(* IEC 61131-3 sources: daoli-st-library/DL_Motion (part 25) *)

(* ---- FB_DL_ToolChangerSeq.st ---- *)
(*
    FB_DL_ToolChangerSeq —— 换刀机构顺控（刀位校验 → 取刀 → 换刀 → 旧刀回库 → 到位确认）
    ------------------------------------------------------------------
    组件名称  : FB_DL_ToolChangerSeq
    分类      : DL_Motion / ToolChange
    前缀      : FB_DL_
    版本      : 1.0.0
    溯源      : 借鉴组织 —— T2-6 Rockwell AOI（矩阵行 166，伺服外围件方向）
                + 次源 t1-9 国产机床 FB 手册公开功能清单（换刀必有反馈对与
                互锁为公开工程惯例）；clean-room 声明 —— 状态机 / 码位 /
                时序 100% 自有，零代码行复制，无闭源参考。
    平台      : 纯 IEC 61131-3（ENUM + CASE + TON / R_TRIG），CODESYS 3.5 /
                TwinCAT 3 / InoProShop / Machine Expert 通用
    作者      : 道莅代码库 · PLC编程专家（R72 构建轮 · 批 4 · 序号 10）
    ------------------------------------------------------------------
    功能说明  : 换刀机构「命令 - 反馈 - 确认」编排：eIdle → eSelect（刀位
                校验 / 映射，发刀位指令，等刀库对位与机械手原位）→ ePick
                （机械手取刀，正向反馈对）→ eSwap（主轴换刀，bSpindleFree
                互锁迁入，反向反馈对）→ eReturn（旧刀回库，回原位反馈）→
                eDone（bToolDone 单拍脉冲）→ eIdle。每执行相带独立超时
                （单 TON 实例，PT = tActTimeout，相驻留即 IN，R145 相级
                看门狗口径），超时 → eFault + 锁存码。
                受理语义（同拍竞态闸，R279）：换刀受理只看 uToolReq **值
                变更沿**的迁入沿锁存副本 _uReqLatch，运行中禁跨拍双判——
                运行中刀位号变更被忽略（沿已被消费），须再次变更刀位号
                （或先归 0）才重新受理；同值重发须先归 0 或变更刀位号
                （接口契约声明，无执行沿引脚的替代口径）。
                安全语义：
                ① eSwap 为安全相，迁入必带全量闸位复检（bSpindleFree +
                   NOT _bFault，R274）；
                ② 换刀中途 bSpindleFree 撤销 → **保持相 + 信息提示，不中断
                   不回退**（防半程掉刀，安全侧声明；继续完成换刀比半程
                   悬臂更安全）；
                ③ 失能 / 故障 → 全输出清零 + 状态回 eIdle（停机相输出清零，
                   R57）；失能不清故障锁存（操作态非复位），复位沿才解除；
                ④ uToolReq = 0 或 > nToolCount → 拒收 + 信息码，不发任何
                   指令；nToolCount = 1（单刀库退化）→ 信息级直接
                   eSelect→ePick（跳过刀库对位等待）。
    错误码    : 16#0004_08B0 刀位请求越域（0 或 > nToolCount），已拒收不发
                            指令 —— 信息级，不置 bError（R45）
                16#0004_08B1 单刀库退化（nToolCount = 1），eSelect 直接转
                            ePick —— 信息级，不置 bError
                16#0004_08B2 执行相超时（任一执行相驻留超 tActTimeout），
                            锁存至复位沿 —— 故障级
                16#0004_08B3 换刀相主轴互锁撤销（bSpindleFree 于 eSwap 内
                            为 FALSE），保持相照走 —— 信息级，不置 bError
                16#0004_08B4 组态非法（nToolCount = 0 / tActTimeout 非正），
                            锁存至复位沿 —— 故障级
                加码反证句（R90）：08B2 / 08B4 输出同为 eFault + bError，
                但 08B4 在 eIdle 即锁存（无执行史）、08B2 必有执行相驻留史
                （eState 轨迹可证），成因互斥不可互换观测；08B0 / 08B1 /
                08B3 各有独立触发事件（拒收沿 / 组态相 / 互锁撤销拍），
                不由现有输出组合还原，故各立一码。
    码位总账  : 16#0004_08B0 用 ｜ 16#0004_08B1 用 ｜ 16#0004_08B2 用 ｜
                16#0004_08B3 用 ｜ 16#0004_08B4 用
                （08A6 / 08A7 已由 FB_DL_TurretToolSelect 占用，本件不占）
    边界与披露: 一 R_TRIG（rtReq / rtReset）与 TON（tonAct）每拍**无条件
                   调用**（规则 ⑦）；tonAct IN = 执行相驻留判据显式变量
                   （R145 看门狗使能只用相驻留，不叠业务条件补集）；超时
                   判定在 CASE 之后（本拍完成事件优先，R275 同拍竞态口径），
                   超时有一拍检测延迟（声明口径）；
                二 零全局变量、零 VAR_EXTERNAL、零物理地址；
                三 归属 Ownership：E_DL_ToolChangePhase 属主为本文件（全库
                   唯一定义，R264），引用件只引用不重声明；
                四 状态机 ENUM + CASE 必带 ELSE 兜底（非法枚举值 → eFault
                   锁存）；段 5b 统一故障迁入闸（R274 迁入完备性）；
                五 反馈引脚语义声明：bToolHome = 所选刀位对位取刀口、
                   bArmHome = 机械手原位、bArmFwd = 机械臂正向到位、
                   bArmBack = 机械臂反向到位，均引脚注入，本件不发轴指令；
                六 分工声明：FB_DL_TurretToolSelect（刀塔分度就近选刀解算，
                   无机械手取放编排）、FB_DL_ToolLifeBudget（寿命记账）——
                   本件只管换刀机构「命令 - 反馈 - 确认」时序编排，刀位
                   就近解算归刀塔件、寿命记账归记账件，互引不互代；
                七 依赖声明：仅 Standard.library（TON / R_TRIG），零厂商
                   方言；
                八 复位沿作用域（R311 逐项声明）：清故障锁存 + 清锁存码 +
                   迁 eIdle + 清 _uReqPrev（强制下次刀位值变更沿可受理），
                   **不清**周期计数类（本件无）与 _uReqLatch（回 Idle 后由
                   下次受理沿重写）。
    验收向量  : V1 正常换刀（uToolReq = 3，nToolCount = 8，反馈按时序到）
                → eState 轨迹 eIdle→eSelect→ePick→eSwap→eReturn→eDone→
                eIdle，bToolDone 单拍，eFault 不出现；
                V2 uToolReq = 0 → 08B0 拒收不发指令；V3 nToolCount = 1 →
                08B1 + eSelect 直转 ePick；V4 eSwap 中 bSpindleFree 撤销
                → 保持相照走 + 08B3；V5 任一执行相超时 → 08B2 锁存 +
                eFault + 输出清零；V6 复位沿 → 解锁回 eIdle；
                V7 nToolCount = 0 → 08B4 锁存；V8 失能 → 输出清零 +
                eIdle，锁存保留。
                算法已证（脚本）：未跑 ｜ 编译器已证（三平台）：未跑
    修订记录  : 2026-11-23 v1.0.0 首次入库（R72 构建轮 · 批 4 · 序号 10）
*)
TYPE E_DL_ToolChangePhase :
(
    eIdle   := 0,                          // 空闲：等刀位请求值变更沿 / idle, waiting for a tool request change edge
    eSelect := 10,                         // 刀位校验：发刀位指令，等刀库对位与机械手原位 / select, issue the tool command
    ePick   := 20,                         // 取刀：机械臂正向，等正向到位 / pick, the arm forward to the magazine
    eSwap   := 30,                         // 换刀：主轴互锁迁入，机械臂反向 / swap, gated by the spindle free interlock
    eReturn := 40,                         // 旧刀回库：机械臂正向回原位 / return, the old tool back to the magazine
    eDone   := 50,                         // 完成：bToolDone 单拍脉冲相 / done, the one shot pulse phase
    eFault  := 60                          // 故障：锁存待复位 / fault, latched until the reset
);
END_TYPE

FUNCTION_BLOCK FB_DL_ToolChangerSeq
VAR_INPUT
    uToolReq     : UINT := 0;              (* 目标刀位请求，[刀位]，1 起计，0 或越容量拒收 / the requested tool number, refused when zero or over capacity *)
    nToolCount   : UINT := 8;              (* 刀库容量组态，[刀位]，禁 0 / the magazine tool count, must not be zero *)
    bToolHome    : BOOL := FALSE;          (* 所选刀位对位反馈，[标志]，引脚注入 / the tool position aligned feedback *)
    bArmHome     : BOOL := FALSE;          (* 机械手原位反馈，[标志]，引脚注入 / the arm home feedback *)
    bArmFwd      : BOOL := FALSE;          (* 机械臂正向到位反馈，[标志]，引脚注入 / the arm forward in position feedback *)
    bArmBack     : BOOL := FALSE;          (* 机械臂反向到位反馈，[标志]，引脚注入 / the arm backward in position feedback *)
    bSpindleFree : BOOL := FALSE;          (* 主轴可换刀互锁，[标志]，eSwap 迁入与驻留判据 / the spindle free interlock *)
    tActTimeout  : TIME := T#10S;          (* 执行相超时，[ms]，禁非正 / the action phase timeout *)
    bEn          : BOOL := FALSE;          (* 使能，[标志]，FALSE 输出清零回 eIdle（锁存保留）/ the enable *)
    bReset       : BOOL := FALSE;          (* 故障复位，[标志]，上升沿唯一解除 / the fault reset *)
END_VAR
VAR_OUTPUT
    uToolSelCmd : UINT := 0;               (* 刀位指令出口，[刀位]，空闲 / 失能 / 故障为 0 / the tool command outlet *)
    bArmFwdCmd  : BOOL := FALSE;           (* 机械臂正向指令出口，[标志] / the arm forward command outlet *)
    bArmBackCmd : BOOL := FALSE;           (* 机械臂反向指令出口，[标志] / the arm backward command outlet *)
    bToolDone   : BOOL := FALSE;           (* 换刀完成单拍脉冲（R24 口径，内部 _bDone 两段式映射）/ the tool done one shot pulse *)
    eState      : E_DL_ToolChangePhase := E_DL_ToolChangePhase.eIdle; // 主状态机当前态 [状态] / the current state
    bError      : BOOL := FALSE;           (* 故障标志，与锁存同源（R191）/ the fault flag from the latch *)
    nErrCode    : UDINT := 16#0000_0000;   (* 错误码，0 = 正常，故障锁存回放（R187）/ the error id *)
END_VAR
VAR
    _bInit     : BOOL := FALSE;            (* 首拍初始化标志（R310）/ the first scan flag *)
    _eState    : E_DL_ToolChangePhase := E_DL_ToolChangePhase.eIdle; // 内部状态寄存器 / the internal state register
    _bFault    : BOOL := FALSE;            (* 故障锁存副本，仅复位沿解除 / the fault latch copy *)
    _nCodeLatch: UDINT := 0;               (* 锁存成因码，故障期回放 / the latched cause code *)
    _uReqLatch : UINT := 0;                (* 受理沿锁存刀位副本（同拍竞态闸，R279）/ the latched tool request copy *)
    _uReqPrev  : UINT := 0;                (* 请求值上一拍快照（值变更沿判据，主体末行刷新，R46）/ the previous request snapshot *)
    _uSelCmd   : UINT := 0;                (* 刀位指令内部副本 / the internal tool command copy *)
    _bFwdCmd   : BOOL := FALSE;            (* 正向指令内部副本 / the internal forward command *)
    _bBackCmd  : BOOL := FALSE;            (* 反向指令内部副本 / the internal backward command *)
    _bDone     : BOOL := FALSE;            (* 完成单拍内部位（段 1 预清，段 5 置位，统一出口映射）/ the internal done bit *)
    _bReqRej   : BOOL := FALSE;            (* 请求拒收信息标志（受理沿消费或复位解除）/ the request rejected info flag *)
    _bDegrade  : BOOL := FALSE;            (* 单刀库退化信息标志 / the single tool degrade info flag *)
    _bSpHold   : BOOL := FALSE;            (* 换刀相互锁撤销信息标志（逐拍重算）/ the spindle hold info flag *)
    _bActive   : BOOL := FALSE;            (* 执行相驻留判据（tonAct IN 显式变量）/ the active phase residency flag *)
    rtReq      : R_TRIG;                   (* 刀位请求值变更沿实例（无条件调用）/ the request change edge instance *)
    rtReset    : R_TRIG;                   (* 复位沿实例（无条件调用）/ the reset edge instance *)
    tonAct     : TON;                      (* 执行相看门狗实例（无条件调用，R145 相驻留使能）/ the action watchdog timer *)
END_VAR
VAR CONSTANT
    DL_TCS_CODE_REQ : UDINT := 16#0004_08B0; (* 请求越域信息码 [码] / the request rejected info code *)
    DL_TCS_CODE_ONE : UDINT := 16#0004_08B1; (* 单刀库退化信息码 [码] / the degrade info code *)
    DL_TCS_CODE_TO  : UDINT := 16#0004_08B2; (* 执行相超时故障码 [码] / the timeout fault code *)
    DL_TCS_CODE_SP  : UDINT := 16#0004_08B3; (* 互锁撤销信息码 [码] / the spindle hold info code *)
    DL_TCS_CODE_CFG : UDINT := 16#0004_08B4; (* 组态非法故障码 [码] / the config fault code *)
    DL_TCS_TZERO    : TIME := T#0S;          (* 零时长哨兵 [ms] / the zero duration sentinel *)
    DL_TCS_ZERO     : UDINT := 0;            (* 无符号零哨兵 [码] / the unsigned zero sentinel *)
    DL_TCS_UZERO    : UINT := 0;             (* 刀位零哨兵 [刀位] / the tool zero sentinel *)
    DL_TCS_UONE     : UINT := 1;             (* 刀位下界哨兵 [刀位] / the tool lower bound sentinel *)
END_VAR

// 段 0｜沿检测与看门狗无条件周期调用（规则 ⑦；IN = 相驻留显式变量）/ segment 0, the unconditional edge and watchdog refresh
rtReq(CLK := (uToolReq <> _uReqPrev));     // 请求值变更沿（同值重发不产生沿，契约声明）/ the request change edge
rtReset(CLK := bReset);                    // 复位沿 / the reset edge
_bActive := (_eState = E_DL_ToolChangePhase.eSelect)   // 执行相驻留判据（R145：只看相驻留）/ the active residency flag
         OR (_eState = E_DL_ToolChangePhase.ePick)
         OR (_eState = E_DL_ToolChangePhase.eSwap)
         OR (_eState = E_DL_ToolChangePhase.eReturn);
tonAct(IN := _bActive AND bEn AND (NOT _bFault), PT := tActTimeout); // 看门狗（失能 / 锁存即断计）/ the watchdog

// 段 1｜首拍初始化与单拍位预清（R310 / FB32-1 / R256）/ segment 1, the first scan init and the presets
IF NOT _bInit THEN                         // 首拍一拍 / the first scan
    _bInit := TRUE;                        // 置首拍标志 / raise the first scan flag
    _bFault := FALSE;                      // 故障锁存显式清零 / clear the fault latch explicitly
    _eState := E_DL_ToolChangePhase.eIdle; // 状态显式落空闲 / place the state to idle
END_IF
_bDone   := FALSE;                         // 完成单拍预清零（置位在段 5 eDone 相）/ preset the done bit false
_bSpHold := FALSE;                         // 互锁撤销标志预清零（eSwap 相逐拍重算）/ preset the hold flag false
_bDegrade := (nToolCount = DL_TCS_UONE) AND _bActive; // 退化信息逐拍重算（执行相驻留内才发码，信息级每拍重算口径 R187）/ the degrade flag recomputed

// 段 2｜复位沿（作用域声明见头注释边界八，R311）/ segment 2, the reset edge with the declared scope
IF rtReset.Q THEN                          // 复位上升沿 / the reset rising edge
    _bFault := FALSE;                      // 清故障锁存（唯一人工解除边，恒可达 R152 自证）/ clear the fault latch
    _nCodeLatch := DL_TCS_ZERO;            // 清锁存码 / clear the latched code
    _eState := E_DL_ToolChangePhase.eIdle; // 迁回空闲 / back to idle
    _uReqPrev := DL_TCS_UZERO;             // 清请求快照（强制下次值变更沿可受理）/ clear the request snapshot
    _bReqRej := FALSE;                     // 清拒收信息标志（复位沿清除边）/ clear the reject flag
END_IF

// 段 3｜组态闸：容量为 0 或超时非正 → 锁存（首次成因，R189）/ segment 3, the configuration gate
IF (NOT _bFault) AND ((nToolCount = DL_TCS_UZERO) OR (tActTimeout <= DL_TCS_TZERO)) THEN // 组态非法命中 / a configuration fault hit
    _bFault := TRUE;                       // 置锁存 / latch the fault
    _nCodeLatch := DL_TCS_CODE_CFG;        // 登记组态码 / register the config code
END_IF

// 段 4｜主状态机（ENUM + CASE，ELSE 兜底；完成事件先于超时判定消化，R275）/ segment 4, the main state machine
CASE _eState OF

    E_DL_ToolChangePhase.eIdle:            // 空闲相 / the idle phase
        _uSelCmd := DL_TCS_UZERO;          // 停机相输出清零（R57）/ zero the command in idle
        _bFwdCmd := FALSE;                 // 指令清零 / clear the commands
        _bBackCmd := FALSE;                // 指令清零 / clear the commands
        IF rtReq.Q AND bEn AND (NOT _bFault) THEN // 受理沿 + 全量闸位复检（R274）/ the accept edge with the gate recheck
            IF (uToolReq >= DL_TCS_UONE) AND (uToolReq <= nToolCount) THEN // 刀位校验（1 起计）/ the tool validation
                _uReqLatch := uToolReq;    // 受理沿锁存副本（R279 禁跨拍双判）/ latch the request copy
                _uSelCmd := _uReqLatch;    // 发刀位指令 / issue the tool command
                _bReqRej := FALSE;         // 受理沿清除旧拒收标志 / clear the old reject flag on accept
                _eState := E_DL_ToolChangePhase.eSelect; // 迁入校验相 / enter the select phase
            ELSE                           // 越域请求拒收（不发任何指令）/ the out of domain request rejected
                _bReqRej := TRUE;          // 置拒收信息标志 / raise the reject flag
            END_IF
        END_IF

    E_DL_ToolChangePhase.eSelect:          // 刀位校验相：等刀库对位与机械手原位 / the select phase
        IF nToolCount = DL_TCS_UONE THEN   // 单刀库退化：跳过对位等待（信息级）/ the single tool degrade
            _bDegrade := TRUE;             // 置退化信息标志 / raise the degrade flag
            _eState := E_DL_ToolChangePhase.ePick; // 直转取刀相 / straight to the pick phase
        ELSIF bToolHome AND bArmHome THEN  // 刀库对位且机械手原位 / the magazine aligned and the arm home
            _eState := E_DL_ToolChangePhase.ePick; // 迁入取刀相 / enter the pick phase
        END_IF

    E_DL_ToolChangePhase.ePick:            // 取刀相：机械臂正向 / the pick phase
        _bFwdCmd := TRUE;                  // 正向指令 / the forward command
        IF bArmFwd AND bSpindleFree AND (NOT _bFault) THEN // 正向到位 + 安全相迁入全量闸位复检（R274）/ the in position with the full gate recheck
            _eState := E_DL_ToolChangePhase.eSwap; // 迁入换刀相 / enter the swap phase
        END_IF                             // 到位但主轴未自由：驻留等待（超时看门狗兜底）/ hold until free

    E_DL_ToolChangePhase.eSwap:            // 换刀相：机械臂反向（互锁撤销保持照走，安全侧声明）/ the swap phase
        _bFwdCmd := FALSE;                 // 撤正向指令 / drop the forward command
        _bBackCmd := TRUE;                 // 反向指令 / the backward command
        _bSpHold := NOT bSpindleFree;      // 互锁撤销逐拍重算（保持相 + 提示，不中断不回退）/ the hold flag recomputed
        IF bArmBack THEN                   // 反向到位 / the backward in position
            _eState := E_DL_ToolChangePhase.eReturn; // 迁入回库相 / enter the return phase
        END_IF

    E_DL_ToolChangePhase.eReturn:          // 旧刀回库相：机械臂正向回原位 / the return phase
        _bBackCmd := FALSE;                // 撤反向指令 / drop the backward command
        _bFwdCmd := TRUE;                  // 正向指令（回库动作）/ the forward command
        IF bArmHome THEN                   // 机械手回原位（旧刀入库确认）/ the arm back home
            _eState := E_DL_ToolChangePhase.eDone; // 迁入完成相 / enter the done phase
        END_IF

    E_DL_ToolChangePhase.eDone:            // 完成相：单拍脉冲（两段式，FB33-1）/ the done phase
        _bDone := TRUE;                    // 置完成单拍内部位 / raise the internal done bit
        _uSelCmd := DL_TCS_UZERO;          // 指令清零 / clear the command
        _bFwdCmd := FALSE;                 // 指令清零 / clear the commands
        _bBackCmd := FALSE;                // 指令清零 / clear the commands
        _eState := E_DL_ToolChangePhase.eIdle; // 迁回空闲（脉冲次拍由段 1 预清撤销，R129 两拍口径）/ back to idle

    E_DL_ToolChangePhase.eFault:           // 故障相：等复位沿（解除可达）/ the fault phase until the reset
        IF NOT _bFault THEN                // 锁存已清才迁出 / the exit after the latch cleared
            _eState := E_DL_ToolChangePhase.eIdle; // 迁回空闲 / back to idle
        END_IF

    ELSE                                   // 非法枚举值拦截 / the illegal enumeration guard
        _eState := E_DL_ToolChangePhase.eFault; // 落故障相 / force to the fault phase
        _bFault := TRUE;                   // 置锁存 / latch the fault
        _nCodeLatch := DL_TCS_CODE_CFG;    // 复用组态码（R90 反证：非法枚举不可达无独立观测需求）/ reuse the config code

END_CASE

// 段 4b｜故障统一迁入闸（置于状态机之后，R274 迁入完备性）/ segment 4b, the unified fault entry gate
IF _bFault AND (_eState <> E_DL_ToolChangePhase.eFault) THEN // 已锁存但不在故障相 / latched but not in the fault phase
    _eState := E_DL_ToolChangePhase.eFault; // 任何相检出故障一律落故障相 / any phase with a latch lands in the fault phase
END_IF

// 段 5｜执行相超时判定（CASE 之后：本拍完成事件已优先消化，R275；超时有一拍
//        检测延迟，声明口径；驻留判据按 CASE 后现值重取，完成迁移即取消超时）/
//        segment 5, the phase timeout verdict with the post CASE residency
IF ((_eState = E_DL_ToolChangePhase.eSelect) OR (_eState = E_DL_ToolChangePhase.ePick)
    OR (_eState = E_DL_ToolChangePhase.eSwap) OR (_eState = E_DL_ToolChangePhase.eReturn))
    AND tonAct.Q THEN                      // 相驻留（现值）且看门狗到时 / the residency with the watchdog expired
    IF NOT _bFault THEN                    // 未锁存才登记超时成因 / register the timeout cause only while not latched
        _bFault := TRUE;                   // 置锁存 / latch the fault
        _nCodeLatch := DL_TCS_CODE_TO;     // 登记超时码 / register the timeout code
    END_IF
END_IF

// 段 6｜失能路径：停机相输出清零 + 回 eIdle（锁存保留，操作态非复位，R57/R191 声明）/ segment 6, the disable path
IF NOT bEn THEN                            // 失能 / disabled
    _eState := E_DL_ToolChangePhase.eIdle; // 状态回空闲 / back to idle
    _uSelCmd := DL_TCS_UZERO;              // 输出清零 / zero the outlets
    _bFwdCmd := FALSE;                     // 指令清零 / clear the commands
    _bBackCmd := FALSE;                    // 指令清零 / clear the commands
    _bReqRej := FALSE;                     // 清拒收信息标志（失能清除边）/ clear the reject flag
END_IF

// 段 7｜统一出口（内部副本单点映射；信息级码优先级：拒收 > 互锁撤销 > 退化，声明口径）/ segment 7, the unified outlet
uToolSelCmd := _uSelCmd;                   // 刀位指令出口 / the tool command outlet
bArmFwdCmd := _bFwdCmd;                    // 正向指令出口 / the forward command outlet
bArmBackCmd := _bBackCmd;                  // 反向指令出口 / the backward command outlet
bToolDone := _bDone;                       // 完成单拍出口（统一出口映射，R189 两段式）/ the done pulse outlet
eState := _eState;                         // 状态出口 / the state outlet
bError := _bFault;                         // 故障标志与锁存同源 / the fault flag from the latch
IF _bFault THEN                            // 故障锁存回放（R187）/ the latched replay
    nErrCode := _nCodeLatch;               // 回放锁存码 / replay the latched code
ELSIF _bReqRej THEN                        // 拒收信息级 / the rejected request
    nErrCode := DL_TCS_CODE_REQ;           // 信息级：请求越域拒收 / info level
ELSIF _bSpHold THEN                        // 互锁撤销信息级 / the spindle hold
    nErrCode := DL_TCS_CODE_SP;            // 信息级：保持相提示 / info level
ELSIF _bDegrade THEN                       // 退化信息级 / the degrade
    nErrCode := DL_TCS_CODE_ONE;           // 信息级：单刀库退化 / info level
ELSE                                       // 无事件 / no event
    nErrCode := DL_TCS_ZERO;               // 正常 / ok
END_IF

// 段 8｜请求值上一拍快照（主体末行无条件刷新，R46 末拍快照口径）/ segment 8, the request snapshot at the body end
_uReqPrev := uToolReq;                     // 末拍快照 / the end of body snapshot
END_FUNCTION_BLOCK

(* ---- FB_DL_TorqueLimitControl.st ---- *)
(*==============================================================================
 * 组件名称 (Component)  : FB_DL_TorqueLimitControl
 * 所属子库 (Sublibrary) : DL_Motion
 * 当前版本 (Version)    : 1.0.0
 * 组件分类 (Category)   : 功能块（FUNCTION_BLOCK）· 压装与力矩族 · 力矩达限压装判定
 * 兼容性   (Platform)   : CODESYS 3.5 / TwinCAT 3 / 汇川 InoProShop / Schneider
 *                         Machine Expert；仅依赖 Standard.library
 *                         （TON / R_TRIG / LIMIT / MIN / MAX / ABS），零厂商方言
 * 接口依赖 (Depends)    : I_DL_MotionAxis / E_DL_AxisState（既有契约，Round 05，零修改）
 * 功能描述 (Function)   : 力矩达限压装判定（「运行到固定挡块」语义的 clean-room 独立
 *                         实现）。流程为 接近 → 慢速压装 → 力矩达限判定 → 达限保持
 *                         → 位移窗口合格判定 → 释放归位。严格区分「设备异常」（未达
 *                         限超时、力矩信号无效、释放超时）与「工件不合格」（到位但
 *                         位移越窗），前者进故障锁存，后者只出判定结果与方向提示。
 * 设计要点 (Key notes)  :
 *   ① 达限判据三源等价（驱动器力矩限制激活 / 实际力矩达阈值 / 驱动器到达挡块反馈），
 *      三者任一成立即判达限，现场按可用信号接入，未接线引脚保持 FALSE 即可。
 *   ② 位移窗判定只在「达限瞬间位置」上做一次锁存判定，判定结果全程保持，避免释放
 *      段位置回退污染结论。
 *   ③ 判定输出先清后置，出口断言「合格与不合格不同时为真」，不合格优先。
 *   ④ 单拍脉冲 bDone 采用「进入态置位、下一拍开头复位」的闭环生命周期，不在同一
 *      扫描内自我清除（单拍标志生命周期三律）。
 *   ⑤ 本块只做判定与流程编排：力矩限幅本身由驱动器参数承担，软件力矩限制不是安全
 *      功能，机械限位与安全回路仍是最终边界。
 * 开源溯源 (Origin)     : 原创实现，clean-room。语义来源为某工业自动化厂商官方支持
 *                         文档的公开页面「转矩限幅及固定停止点检测」（两种模式分离、
 *                         达限状态输出）、公开技术知识库页面（挡块力矩 / 位置检测窗
 *                         / 到达挡块最长时限的参数域）（来源编号 RAW_NOTES S-4）。
 *                         「借鉴对象的许可说明」：上述对象为该厂商免费使用但闭源
 *                         版权的官方文档与公开技术文章，属「可免费查阅、仅借鉴参数
 *                         域与状态语义」类别；本实现未复制任何示例程序、源码或组态
 *                         数据，状态机、判定逻辑、故障码 100% 自有设计；亦不实现
 *                         厂商的力矩限幅指令本身（本库接口无扭矩域，扭矩经引脚注入）。
 * 验收向量 (Acceptance) :
 *   V1 正常压装：达限位置 20.5 mm、位移窗 20.0~21.0 → bJudgeOk 为 TRUE；
 *   V2 压到 19.5 mm（低于窗下限）→ bJudgeNg 为 TRUE 且出信息级 0163；
 *   V3 压到 21.5 mm（高于窗上限）→ bJudgeNg 为 TRUE 且出信息级 0164；
 *   V4 压装段 10 s 未达限 → 锁存 0282（工件过软 / 未到位 / 信号失效）；
 *   V5 终点不超过起点 → 启动沿锁存 0280（方向组态错误）；
 *   V6 位移窗写反（低 21 / 高 20）→ 对调自修复 + 信息级 0160，判定仍有效；
 *   V7 中途 bAbort → 立即受控停止退回，判定输出清零且不置不合格；
 *   V8 fActTorque 为非有限值 → 锁存 0283（判定不可信）；
 *   V9 运行中途插入跟踪脉冲 bTrack：清判定与锁存、退回 eIdle（公约 0.1）。
 * 已知限制 (Limits)     :
 *   ① 力矩与达限状态由驱动适配层经引脚注入（轴接口无扭矩域），本块不读取驱动器
 *      内部参数；引脚未接时达限判据退化为阈值比较，可能永远等不到达限。
 *   ② 释放目标固定取压装起点（不引入额外释放位引脚），若工艺需要退到更远的安全
 *      位，请在上层压制完成后追加一条定位指令。
 *   ③ 本块为判定层与流程编排层，不构成 ISO 13849 / IEC 62061 认证安全功能。
 * 规格偏离 (Deviation)  :
 *   ① 依公约 0.1 增补 bTrack 输入引脚（首扫 / 跟踪范式强制项）。
 *   ② eRelease 超时按故障级 0281 处理并进入 eFault，而非留在 eDone 带码：
 *      规格仅写「超时置故障 0281，不静默」，本块取严格处置，避免上层误判合格。
 *   ③ 速度 / 力矩参数非正或非有限值时回默认值（与库内其他运动件口径一致），
 *      不在启动沿判故障；力矩阈值超额定只提示不阻断（依规格 0161 语义）。
 *   ④ 使能撤除时补发一次停止请求（安全保守处置）。
 * 红线自检 (Redline)    :
 *   R1 零全局符号区访问 ✓（无全局变量表访问、无外部变量声明）
 *   R2 零物理地址直写 ✓（无输入输出通道地址记号）
 *   R3 纯 IEC 61131-3 ✓（仅 TON / R_TRIG / LIMIT / MIN / MAX / ABS）
 *   R4 防除零 / 防越界 / 浮点容差 ✓（无除法、浮点比较全用容差、无数组索引）
 *   R5 声明行 100% 中英双语同行注释 ✓
 *   R6 ENUM + CASE 且 CASE 含 ELSE 兜底 ✓
 *   R7 定时器与边沿实例无条件周期刷新 ✓；单拍标志 bDone 置位于本次进入、复位于
 *      下一拍开头，同一周期闭环，无跨周期残留 ✓
 *   POU 终结符成对 ✓（FUNCTION_BLOCK ↔ END_FUNCTION_BLOCK，末行即终结符；
 *   TYPE ↔ END_TYPE 成对）
 * 故障码表 (Error codes):
 *   16#0004_0160【信息级】位移窗上下限对调自修复；
 *   16#0004_0161【信息级】达限力矩超额定（机械风险提示）；
 *   16#0004_0162【信息级】压装速度高于接近速度（工艺反常）；
 *   16#0004_0163【信息级】到位但位移低于窗下限（压浅，判定方向提示）；
 *   16#0004_0164【信息级】到位但位移高于窗上限（压深，判定方向提示）；
 *   16#0004_0280【故障级】压装行程组态非法（终点不大于起点 / 位置非有限值），锁存；
 *   16#0004_0281【故障级】释放超时，锁存；
 *   16#0004_0282【故障级】压装超时未达限，锁存；
 *   16#0004_0283【故障级】力矩信号非有限值，锁存；
 *   16#0004_0284【故障级】轴指令被拒 / 轴故障，锁存；
 *   16#0004_0296【故障级】非法状态兜底（本块专用，不与其他块共用）。
 *   信息级码只进 uErrorId；bError 为派生式仅反映 eFault 态。
 * 修订历史 (Revision)   :
 *   2026-11-15  v1.0.0  首版入库（Round 08 · DL_Motion 压装与力矩族开族件）
 *============================================================================*)

(*-----------------------------------------------------------------------------
 * 调用示例 (Instance guide)：
 *   fbPress.iAxis := fbPressAxis;                  // 压装轴实例注入
 *   fbPress(bEnable := TRUE, bStart := bStartPress,
 *           fPressStartPos := 10.0, fPressEndPos := 30.0,
 *           fPosWindowLow := 20.0, fPosWindowHigh := 21.0,
 *           fTorqueLimit := 30.0,
 *           fApproachVel := 50.0, fPressVel := 5.0, fAcc := 200.0,
 *           tClampTime := T#300MS, tPressTimeout := T#10S,
 *           fActTorque := fDriveTorque,
 *           bTorqueLimitActive := bDriveInLimitation);
 *   IF fbPress.bDone THEN
 *       bResultOk := fbPress.bJudgeOk;             // 只在 bDone 单拍内取结果
 *   END_IF
 *   注：驱动器侧的力矩限幅（如力矩上限参数族）与「到达挡块」功能必须先行组态，
 *       本块只消费其状态反馈，不代替驱动器限幅。
 *----------------------------------------------------------------------------*)

(*-----------------------------------------------------------------------------
 * 常见误用与现场提示 (Field notes)：
 *   1 压装速度经验值取接近速度的 1/10 左右；压装快于接近速度时本块只提示
 *      （信息级 0162），不会拒绝执行，但冲击会损伤工件与压头。
 *   2 位移窗必须按「达限瞬间位置」组态，而不是按「起点到终点」的行程；窗上下限
 *      填反会被自动对调并提示，但仍建议在配方里改对。
 *   3 力矩阈值填超过额定值（>100）只提示不阻断，属于「明知有机械风险仍要压」的
 *      场景；正式产线请把上限压回 100 以内。
 *   4 bAbort 是电平最高优先：任意态给 TRUE 立即受控停止并退回空闲，判定结果清零，
 *      不会把中途中止误判为不合格工件。
 *   5 bDone 只维持一个扫描周期，上层必须在本拍内取 bJudgeOk / bJudgeNg 并存到
 *      自己的结果寄存器里；跨拍读判定请读 bJudgeOk / bJudgeNg（这两者在 eDone
 *      期间保持）。
 *----------------------------------------------------------------------------*)

(*-----------------------------------------------------------------------------
 * 枚举: E_DL_PressState（归属 DL_Motion，与本功能块同文件发布）
 * 含义: 力矩达限压装流程状态机，编号间隔 10 预留扩展位。
 *----------------------------------------------------------------------------*)
{attribute 'strict'}
{attribute 'qualified_only'}
TYPE E_DL_PressState :
(
    eIdle     := 0,    // 空闲：未启动，输出清零 / Idle: not started, outputs cleared
    eApproach := 10,   // 接近：以接近速度走向压装起点 / Approach: move to press start at approach speed
    ePress    := 20,   // 压装：以压装速度慢速压入，等力矩达限 / Press: slow press until torque limit reached
    eClamp    := 30,   // 达限保持：力矩达限后保位并计时（应力松弛） / Clamp: hold position and time after torque limit
    eRelease  := 40,   // 释放：退回压装起点 / Release: retract to press start position
    eDone     := 50,   // 完成：判定结果有效，等新启动沿 / Done: judgement valid, waiting for new start edge
    eFault    := 99    // 故障锁存：仅 bReset 上升沿可退出 / Fault: latched, only bReset rising edge exits
) UINT;
END_TYPE

FUNCTION_BLOCK FB_DL_TorqueLimitControl
VAR_INPUT
    bEnable            : BOOL := FALSE;     // 总使能（Enable），FALSE=中止流程并清输出，电平语义
    bStart             : BOOL := FALSE;     // 启动压装周期（Start），上升沿受理，仅 eIdle / eDone 受理
    bAbort             : BOOL := FALSE;     // 中止（Abort），电平最高优先，立即受控停止并退回空闲
    bReset             : BOOL := FALSE;     // 复位故障与判定结果（Reset），上升沿受理
    bTrack             : BOOL := FALSE;     // 内部锁存重同步（Tracking pulse），上升沿清判定与故障并退回 eIdle
    fPressStartPos     : REAL := 0.0;       // 压装起点位置（Press start position）[mm]，接近段目标与释放目标
    fPressEndPos       : REAL := 0.0;       // 压装终点位置（Press end position）[mm]，必须大于起点
    fPosWindowLow      : REAL := 0.0;       // 到位位移窗下限（Position window low）[mm]，窗上下限写反自动对调
    fPosWindowHigh     : REAL := 0.0;       // 到位位移窗上限（Position window high）[mm]
    fTorqueLimit       : REAL := 30.0;      // 达限判定力矩（Torque limit）[% 额定]，域 1..150，>100 仅提示
    fApproachVel       : REAL := 50.0;      // 接近速度（Approach velocity）[mm/s]，域 0.1..1000，非正值回默认
    fPressVel          : REAL := 5.0;       // 压装速度（Press velocity）[mm/s]，域 0.1..100，建议不超接近速度 1/10
    fAcc               : REAL := 200.0;     // 加/减速度（Acceleration）[mm/s²]，域 0.1..100000，非有限值回默认
    tClampTime         : TIME := T#300MS;   // 达限保持时间（Clamp hold time）[ms]，域 T#0S..T#10S
    tPressTimeout      : TIME := T#10S;     // 压装超时（Press timeout）[ms]，域 T#100MS..T#60S
    tReleaseTimeout    : TIME := T#5S;      // 释放超时（Release timeout）[ms]，超时判故障级
    fActTorque         : REAL := 0.0;       // 实际力矩（Actual torque）[% 额定]，由驱动适配层注入
    bTorqueLimitActive : BOOL := FALSE;     // 驱动器力矩限制已激活反馈（Drive in limitation），由适配层注入
    bInClampFeedback   : BOOL := FALSE;     // 驱动器到达固定挡块反馈（Fixed stop reached），可选，未接线保持 FALSE
END_VAR
VAR_OUTPUT
    bJudgeOk           : BOOL := FALSE;     // 判定合格（Judge OK），eDone 内保持
    bJudgeNg           : BOOL := FALSE;     // 判定不合格（Judge NG），eDone 内保持，与合格互斥且优先
    bInClamp           : BOOL := FALSE;     // 已达限压紧（In clamp），eClamp 态为 TRUE
    bBusy              : BOOL := FALSE;     // 周期执行中（Busy），接近 / 压装 / 保持 / 释放四态为 TRUE
    bDone              : BOOL := FALSE;     // 周期结束单拍脉冲（Done pulse），仅进入 eDone 那一拍为 TRUE
    fPosAtClamp        : REAL := 0.0;       // 达限瞬间位置（Position at clamp）[mm]，锁存值
    fTorqueAtClamp     : REAL := 0.0;       // 达限瞬间力矩（Torque at clamp）[% 额定]，锁存值
    bError             : BOOL := FALSE;     // 故障锁存（Error），派生式仅故障级码参与，信息级码不置位
    uErrorId           : UDINT := 0;        // 故障码（Error code），段位 16#0004_xxxx，0=无故障
    nCycleCount        : UDINT := 0;        // 完成周期计数（Cycle counter）[次]，每次进入 eDone 加一
END_VAR
VAR_IN_OUT
    iAxis              : I_DL_MotionAxis;   // 压装轴接口引用（Press axis），由调用方注入实现块实例
END_VAR
VAR
    eState             : E_DL_PressState := E_DL_PressState.eIdle; // 内部状态机步序（Internal state）
    bInit              : BOOL := FALSE;     // 首扫完成标志（First-scan done flag），初值 FALSE，随 bTrack 复位
    bFaultLatch        : BOOL := FALSE;     // 故障锁存标志（Fault latch），仅 bReset 沿或新启动沿解除
    bStopIssued        : BOOL := FALSE;     // 停止已下发标志（Stop issued flag），单发化防重复发令
    bTorqueReached     : BOOL := FALSE;     // 达限标志（Torque limit reached），三源 OR 结果
    bClampTimerBrk     : BOOL := FALSE;     // 保持计时断输入标志（Clamp timer break），时间参数变更时置位
    bPressTimerBrk     : BOOL := FALSE;     // 压装计时断输入标志（Press timer break），时间参数变更时置位
    bRelTimerBrk       : BOOL := FALSE;     // 释放计时断输入标志（Release timer break），时间参数变更时置位
    fWinLowEff         : REAL := 0.0;       // 生效位移窗下限（Effective window low）[mm]，对调后的较小值
    fWinHighEff        : REAL := 0.0;       // 生效位移窗上限（Effective window high）[mm]，对调后的较大值
    fTorqueLimitEff    : REAL := 30.0;      // 生效力矩阈值（Effective torque limit）[% 额定]，已做域钳位
    fApproachEff       : REAL := 50.0;      // 生效接近速度（Effective approach velocity）[mm/s]
    fPressEff          : REAL := 5.0;       // 生效压装速度（Effective press velocity）[mm/s]
    fAccEff            : REAL := 200.0;     // 生效加减速度（Effective acceleration）[mm/s²]
    fPosNow            : REAL := 0.0;      // 轴当前实际位置（Actual position）[mm]
    fTorqueNow         : REAL := 0.0;      // 力矩当前值（Actual torque）[% 额定]，非有限值时按 0 记账
    tClampEff          : TIME := T#300MS;   // 生效保持时间（Effective clamp time）[ms]，负值归零
    tPressEff          : TIME := T#10S;     // 生效压装超时（Effective press timeout）[ms]
    tRelEff            : TIME := T#5S;      // 生效释放超时（Effective release timeout）[ms]
    tClampPrev         : TIME := T#0MS;     // 上拍保持时间（Previous clamp time）[ms]，变更检测基准
    tPressPrev         : TIME := T#0MS;     // 上拍压装超时（Previous press timeout）[ms]，变更检测基准
    tRelPrev           : TIME := T#0MS;     // 上拍释放超时（Previous release timeout）[ms]，变更检测基准
    fbTrigStart        : R_TRIG;            // 启动指令上升沿（Start command rising edge）
    fbTrigReset        : R_TRIG;            // 复位指令上升沿（Reset command rising edge）
    fbTonClamp         : TON;               // 达限保持计时（Clamp hold timer）
    fbTonPressTimeout  : TON;               // 压装超时监控（Press timeout timer）
    fbTonRelTimeout    : TON;               // 释放超时监控（Release timeout timer）
END_VAR
VAR CONSTANT
    DL_PRESS_INF_MAX     : REAL := 1.0E30;  // 有限值判定幅值上限（Finite magnitude bound）[无量纲，按比较量量纲同值使用]
    DL_PRESS_EPS         : REAL := 1.0E-6;  // 浮点判零容差（Float zero tolerance）[无量纲，按比较量量纲同值使用]
    DL_PRESS_POS_BAND    : REAL := 0.05;    // 到位判定带（In-position band）[mm]，位置差小于此值判到位
    DL_PRESS_PAR_FLOOR   : REAL := 1.0E-3;  // 速度/加速度参数下限（Parameter floor）[mm/s 或 mm/s²]
    DL_PRESS_APPR_DEF    : REAL := 50.0;    // 接近速度默认值（Default approach velocity）[mm/s]
    DL_PRESS_PRESS_DEF   : REAL := 5.0;     // 压装速度默认值（Default press velocity）[mm/s]
    DL_PRESS_ACC_DEF     : REAL := 200.0;   // 加速度默认值（Default acceleration）[mm/s²]
    DL_PRESS_VEL_MAX     : REAL := 1000.0;  // 接近速度上限（Approach velocity ceiling）[mm/s]，超限钳位
    DL_PRESS_TQ_DEF      : REAL := 30.0;    // 力矩阈值默认值（Default torque limit）[% 额定]
    DL_PRESS_TQ_NOMINAL  : REAL := 100.0;   // 额定力矩（Nominal torque）[% 额定]，超此值仅提示
    DL_PRESS_TQ_MAX      : REAL := 150.0;   // 力矩阈值上限（Torque limit ceiling）[% 额定]，超限钳位
    DL_PRESS_ZERO_TIME   : TIME := T#0S;    // 零时间字面量（Zero time literal）[ms]，用于时间下限比较
END_VAR

// 段 1｜边沿实例无条件周期刷新（红线 R7：严禁置于 IF / CASE 分支内）
fbTrigStart(CLK := bStart);
fbTrigReset(CLK := bReset);

// 段 2｜出口默认赋值（公约 0.9：早退路径输出必须确定）；bDone 在此复位 = 单拍闭环
bBusy      := FALSE;
bInClamp   := FALSE;
bDone      := FALSE;
bError     := (eState = E_DL_PressState.eFault);

// 段 3｜接口引用有效性防御：未注入轴引用则清输出退出
IF iAxis = 0 THEN
    RETURN;
END_IF

// 段 4｜参数防御：速度 / 加速度 / 力矩阈值非正或非有限值回默认，位移窗写反自动对调
IF (fApproachVel <> fApproachVel) OR (ABS(fApproachVel) > DL_PRESS_INF_MAX)
   OR (fApproachVel < DL_PRESS_PAR_FLOOR) THEN
    fApproachEff := DL_PRESS_APPR_DEF;                    // 接近速度非法 → 默认
ELSE
    fApproachEff := MIN(fApproachVel, DL_PRESS_VEL_MAX);   // 合法 → 上限钳位
END_IF

IF (fPressVel <> fPressVel) OR (ABS(fPressVel) > DL_PRESS_INF_MAX)
   OR (fPressVel < DL_PRESS_PAR_FLOOR) THEN
    fPressEff := DL_PRESS_PRESS_DEF;                      // 压装速度非法 → 默认
ELSE
    fPressEff := MIN(fPressVel, fApproachEff);            // 合法 → 不超接近速度（超出部分另出信息码提示）
END_IF

IF (fAcc <> fAcc) OR (ABS(fAcc) > DL_PRESS_INF_MAX) OR (fAcc < DL_PRESS_PAR_FLOOR) THEN
    fAccEff := DL_PRESS_ACC_DEF;
ELSE
    fAccEff := fAcc;
END_IF

IF (fTorqueLimit <> fTorqueLimit) OR (ABS(fTorqueLimit) > DL_PRESS_INF_MAX)
   OR (fTorqueLimit < DL_PRESS_PAR_FLOOR) THEN
    fTorqueLimitEff := DL_PRESS_TQ_DEF;                   // 力矩阈值非法 → 默认
ELSE
    fTorqueLimitEff := MIN(fTorqueLimit, DL_PRESS_TQ_MAX); // 合法 → 上限钳位 150%
END_IF

fWinLowEff  := fPosWindowLow;
fWinHighEff := fPosWindowHigh;
IF (fWinLowEff <> fWinLowEff) OR (fWinHighEff <> fWinHighEff) THEN
    fWinLowEff  := 0.0;                                   // 非有限值：窗回零，判定必然趋向不合格
    fWinHighEff := 0.0;
ELSIF fWinLowEff > (fWinHighEff - DL_PRESS_EPS) THEN
    fWinLowEff  := fPosWindowHigh;                        // 写反：对调自修复，不静默
    fWinHighEff := fPosWindowLow;
    uErrorId    := 16#0004_0160;                          // 【信息级】位移窗上下限对调自修复
END_IF

// 段 5｜时间参数防御与变更检测（公约 0.6：语义参数变化必须断输入一拍使计时归零）
IF tClampTime < DL_PRESS_ZERO_TIME THEN
    tClampEff := DL_PRESS_ZERO_TIME;
ELSE
    tClampEff := tClampTime;
END_IF
IF tPressTimeout < DL_PRESS_ZERO_TIME THEN
    tPressEff := DL_PRESS_ZERO_TIME;
ELSE
    tPressEff := tPressTimeout;
END_IF
IF tReleaseTimeout < DL_PRESS_ZERO_TIME THEN
    tRelEff := DL_PRESS_ZERO_TIME;
ELSE
    tRelEff := tReleaseTimeout;
END_IF
bClampTimerBrk := (tClampEff <> tClampPrev);
bPressTimerBrk := (tPressEff <> tPressPrev);
bRelTimerBrk   := (tRelEff <> tRelPrev);
tClampPrev     := tClampEff;
tPressPrev     := tPressEff;
tRelPrev       := tRelEff;

// 段 6｜反馈量采集与信号有效性判定
fPosNow := iAxis.fPosition;
IF (fActTorque <> fActTorque) OR (ABS(fActTorque) > DL_PRESS_INF_MAX) THEN
    fTorqueNow  := 0.0;                                   // 力矩信号无效：按零记账，另由状态机置故障级
    bTorqueReached := FALSE;
ELSE
    fTorqueNow  := fActTorque;
    // 达限三源等价：驱动器限制激活 / 实际力矩达阈值 / 到达挡块反馈，任一成立即达限
    bTorqueReached := bTorqueLimitActive OR (fTorqueNow >= fTorqueLimitEff) OR bInClampFeedback;
END_IF

// 段 7｜定时器无条件周期刷新（红线 R7：严禁置于 IF / CASE 分支内）
fbTonClamp(IN := (eState = E_DL_PressState.eClamp) AND (NOT bClampTimerBrk), PT := tClampEff);
fbTonPressTimeout(IN := (eState = E_DL_PressState.ePress) AND (NOT bPressTimerBrk), PT := tPressEff);
fbTonRelTimeout(IN := (eState = E_DL_PressState.eRelease) AND (NOT bRelTimerBrk), PT := tRelEff);

// 段 8｜首扫与跟踪范式（公约 0.1：bTrack OR (NOT bInit) 为唯一判据，禁止反序）
IF bTrack OR (NOT bInit) THEN
    bFaultLatch    := FALSE;
    bStopIssued    := FALSE;
    bJudgeOk       := FALSE;
    bJudgeNg       := FALSE;
    fPosAtClamp    := 0.0;                                // 达限位置锁存清零 [mm]
    fTorqueAtClamp := 0.0;                                // 达限力矩锁存清零 [% 额定]
    eState         := E_DL_PressState.eIdle;
    bInit          := TRUE;                               // 首扫完成后置位（判据恒为 bTrack OR NOT bInit）
END_IF

// 段 9｜总使能撤除：中止流程 + 补发一次停止（安全保守处置）
IF NOT bEnable THEN
    IF (NOT bStopIssued) AND (eState <> E_DL_PressState.eIdle) AND (eState <> E_DL_PressState.eFault) THEN
        iAxis.Stop();                                     // 使能撤除瞬间单发停止
        bStopIssued := TRUE;
    END_IF
    eState     := E_DL_PressState.eIdle;
    bJudgeOk   := FALSE;
    bJudgeNg   := FALSE;
    bInClamp   := FALSE;
END_IF

// 段 10｜中止最高优先：任意运行态立即受控停止并退回空闲（不置不合格，避免误判工件）
IF bAbort AND (eState <> E_DL_PressState.eIdle) AND (eState <> E_DL_PressState.eFault) THEN
    IF NOT bStopIssued THEN
        iAxis.Stop();                                     // 中止单发停止（本拍唯一一次轴调用）
        bStopIssued := TRUE;
    END_IF
    bJudgeOk   := FALSE;
    bJudgeNg   := FALSE;
    bInClamp   := FALSE;
    bBusy      := FALSE;
    eState     := E_DL_PressState.eIdle;
END_IF

// 段 11｜事件码管理（公约 0.7 / R15）：锁存码仅在解除路径清，瞬时码逐拍重算
IF NOT bFaultLatch THEN
    uErrorId := 0;
END_IF

// 段 11.5｜轴位置非有限值拦截（反馈不可信时不得继续判定，按轴异常处置）
IF (fPosNow <> fPosNow) OR (ABS(fPosNow) > DL_PRESS_INF_MAX) THEN
    IF (eState <> E_DL_PressState.eIdle) AND (eState <> E_DL_PressState.eFault) THEN
        bFaultLatch := TRUE;
        uErrorId    := 16#0004_0284;                      // 【故障级】轴位置非有限值（按压装轴异常处置）
        eState      := E_DL_PressState.eFault;
    END_IF
END_IF

// 段 12｜主状态机（ENUM + CASE + ELSE 兜底）
CASE eState OF

    E_DL_PressState.eIdle:                                // 空闲：等待启动沿与组态校验
        bBusy    := FALSE;
        bInClamp := FALSE;
        IF fbTrigStart.Q AND bEnable AND (NOT bAbort) THEN
            bFaultLatch := FALSE;                         // 新启动沿：锁存码解除路径（R15）
            bJudgeOk    := FALSE;
            bJudgeNg    := FALSE;
            bStopIssued := FALSE;
            IF (fPressEndPos <> fPressEndPos) OR (fPressStartPos <> fPressStartPos)
               OR (ABS(fPressEndPos) > DL_PRESS_INF_MAX) OR (ABS(fPressStartPos) > DL_PRESS_INF_MAX)
               OR ((fPressEndPos - fPressStartPos) <= DL_PRESS_EPS) THEN
                bFaultLatch := TRUE;
                uErrorId    := 16#0004_0280;              // 【故障级】压装行程组态非法（终点不大于起点 / 位置非有限值）
                eState      := E_DL_PressState.eFault;
            ELSE
                IF fTorqueLimitEff > DL_PRESS_TQ_NOMINAL THEN
                    uErrorId := 16#0004_0161;             // 【信息级】达限力矩超额定（机械风险提示）
                ELSIF fPressVel > fApproachVel THEN
                    uErrorId := 16#0004_0162;             // 【信息级】压装速度高于接近速度（工艺反常）
                END_IF
                fPosAtClamp    := 0.0;
                fTorqueAtClamp := 0.0;
                eState         := E_DL_PressState.eApproach;
            END_IF
        END_IF

    E_DL_PressState.eApproach:                            // 接近：以接近速度走向压装起点
        bBusy := TRUE;
        IF iAxis.bError THEN
            bFaultLatch := TRUE;
            uErrorId    := 16#0004_0284;                  // 【故障级】轴故障
            eState      := E_DL_PressState.eFault;
        ELSIF ABS(fPosNow - fPressStartPos) <= DL_PRESS_POS_BAND THEN
            eState := E_DL_PressState.ePress;             // 到位 → 进入压装段
        ELSE
            IF NOT iAxis.MoveAbsolute(fPos := fPressStartPos, fVel := fApproachEff, fAcc := fAccEff) THEN
                bFaultLatch := TRUE;
                uErrorId    := 16#0004_0284;              // 【故障级】轴指令被拒
                eState      := E_DL_PressState.eFault;
            END_IF
        END_IF

    E_DL_PressState.ePress:                               // 压装：慢速压入，等力矩达限
        bBusy := TRUE;
        IF iAxis.bError THEN
            bFaultLatch := TRUE;
            uErrorId    := 16#0004_0284;                  // 【故障级】轴故障
            eState      := E_DL_PressState.eFault;
        ELSIF (fActTorque <> fActTorque) OR (ABS(fActTorque) > DL_PRESS_INF_MAX) THEN
            bFaultLatch := TRUE;
            uErrorId    := 16#0004_0283;                  // 【故障级】力矩信号非有限值，判定不可信
            eState      := E_DL_PressState.eFault;
        ELSIF bTorqueReached THEN
            fPosAtClamp    := fPosNow;                     // 锁存达限瞬间位置 [mm]
            fTorqueAtClamp := fTorqueNow;                  // 锁存达限瞬间力矩 [% 额定]
            eState         := E_DL_PressState.eClamp;      // 进入达限保持段
        ELSIF fbTonPressTimeout.Q THEN
            bFaultLatch := TRUE;
            uErrorId    := 16#0004_0282;                  // 【故障级】压装超时未达限
            eState      := E_DL_PressState.eFault;
        ELSE
            IF NOT iAxis.MoveAbsolute(fPos := fPressEndPos, fVel := fPressEff, fAcc := fAccEff) THEN
                bFaultLatch := TRUE;
                uErrorId    := 16#0004_0284;              // 【故障级】轴指令被拒
                eState      := E_DL_PressState.eFault;
            END_IF
        END_IF

    E_DL_PressState.eClamp:                               // 达限保持：零速保位并计时
        bBusy    := TRUE;
        bInClamp := TRUE;
        IF iAxis.bError THEN
            bFaultLatch := TRUE;
            uErrorId    := 16#0004_0284;                  // 【故障级】轴故障
            eState      := E_DL_PressState.eFault;
        ELSIF fbTonClamp.Q THEN
            // 保持结束：按达限瞬间位置做位移窗判定（先清后置，不合格优先）
            bJudgeOk   := FALSE;
            bJudgeNg   := FALSE;
            IF (fPosAtClamp >= fWinLowEff) AND (fPosAtClamp <= fWinHighEff) THEN
                bJudgeOk := TRUE;                         // 落在窗内：合格
            ELSE
                bJudgeNg := TRUE;                         // 越窗：不合格
                IF fPosAtClamp < fWinLowEff THEN
                    uErrorId := 16#0004_0163;             // 【信息级】压浅（低于窗下限）
                ELSE
                    uErrorId := 16#0004_0164;             // 【信息级】压深（高于窗上限）
                END_IF
            END_IF
            bInClamp   := FALSE;
            eState     := E_DL_PressState.eRelease;
        ELSE
            IF NOT iAxis.MoveVelocity(fVel := 0.0, fAcc := fAccEff) THEN
                bFaultLatch := TRUE;
                uErrorId    := 16#0004_0284;              // 【故障级】保位指令被拒
                eState      := E_DL_PressState.eFault;
            END_IF
        END_IF

    E_DL_PressState.eRelease:                             // 释放：退回压装起点
        bBusy := TRUE;
        IF iAxis.bError THEN
            bFaultLatch := TRUE;
            uErrorId    := 16#0004_0284;                  // 【故障级】轴故障
            eState      := E_DL_PressState.eFault;
        ELSIF ABS(fPosNow - fPressStartPos) <= DL_PRESS_POS_BAND THEN
            bBusy        := FALSE;
            bDone        := TRUE;                         // 单拍脉冲：本拍置位，下一拍开头复位
            nCycleCount  := nCycleCount + 1;              // 完成周期计数 [次]
            bStopIssued  := FALSE;
            eState       := E_DL_PressState.eDone;
        ELSIF fbTonRelTimeout.Q THEN
            bFaultLatch := TRUE;
            uErrorId    := 16#0004_0281;                  // 【故障级】释放超时（不静默，避免上层误判合格）
            eState      := E_DL_PressState.eFault;
        ELSE
            IF NOT iAxis.MoveAbsolute(fPos := fPressStartPos, fVel := fApproachEff, fAcc := fAccEff) THEN
                bFaultLatch := TRUE;
                uErrorId    := 16#0004_0284;              // 【故障级】轴指令被拒
                eState      := E_DL_PressState.eFault;
            END_IF
        END_IF

    E_DL_PressState.eDone:                                // 完成：判定保持，等新启动沿或复位
        bBusy    := FALSE;
        bInClamp := FALSE;
        IF fbTrigReset.Q THEN
            bJudgeOk   := FALSE;
            bJudgeNg   := FALSE;
            eState     := E_DL_PressState.eIdle;
        ELSIF fbTrigStart.Q AND bEnable AND (NOT bAbort) THEN
            bJudgeOk   := FALSE;                          // 新周期：判定清零后重新压装
            bJudgeNg   := FALSE;
            fPosAtClamp    := 0.0;
            fTorqueAtClamp := 0.0;
            bStopIssued    := FALSE;
            IF (fPressEndPos <> fPressEndPos) OR (fPressStartPos <> fPressStartPos)
               OR ((fPressEndPos - fPressStartPos) <= DL_PRESS_EPS) THEN
                bFaultLatch := TRUE;
                uErrorId    := 16#0004_0280;              // 【故障级】压装行程组态非法
                eState      := E_DL_PressState.eFault;
            ELSE
                eState := E_DL_PressState.eApproach;
            END_IF
        END_IF

    E_DL_PressState.eFault:                               // 故障锁存：仅复位沿可退出
        bBusy      := FALSE;
        bInClamp   := FALSE;
        bStopIssued := FALSE;
        IF fbTrigReset.Q THEN
            bFaultLatch    := FALSE;                      // 唯一解除路径
            uErrorId       := 0;
            bJudgeOk       := FALSE;
            bJudgeNg       := FALSE;
            fPosAtClamp    := 0.0;
            fTorqueAtClamp := 0.0;
            eState         := E_DL_PressState.eIdle;
        END_IF

    ELSE                                                  // 非法状态兜底（本块专用码）
        bFaultLatch := TRUE;
        uErrorId    := 16#0004_0296;                      // 【故障级】非法状态兜底
        bBusy       := FALSE;
        bInClamp    := FALSE;
        eState      := E_DL_PressState.eFault;

END_CASE

// 段 13｜出口映射与判定互斥断言（不合格优先，两者不得同真）
bError   := (eState = E_DL_PressState.eFault);
bInClamp := (eState = E_DL_PressState.eClamp);
bBusy    := (eState = E_DL_PressState.eApproach) OR (eState = E_DL_PressState.ePress)
            OR (eState = E_DL_PressState.eClamp) OR (eState = E_DL_PressState.eRelease);
IF bJudgeOk AND bJudgeNg THEN
    bJudgeOk := FALSE;                                    // 互斥断言：同时为真时按不合格处置
    bJudgeNg := TRUE;
END_IF

END_FUNCTION_BLOCK

(* ---- FB_DL_WinderTensionTaperCalc.st ---- *)
(*==============================================================================
 * 组件名称 (Component)  : FB_DL_WinderTensionTaperCalc
 * 所属子库 (Sublibrary) : DL_Motion ｜ 版本 (Version) : 1.0.0 ｜ 2026-11-23
 * 兼容性   (Platform)   : CODESYS 3.5+ / TwinCAT 3 / 汇川 InoProShop / 施耐德 Machine Expert
 *                         仅依赖 IEC 61131-3 标准（CASE / ABS / MAX / MIN），零厂商私有库
 * 功能描述 (Function)   : 收卷锥度张力计算（分段折线口径）。卷径归一化比例 r =
 *                         (fRollDia − fDiaCore) ÷ (fDiaMax − fDiaCore) ∈ [0,1]，锥度系数 k(r)
 *                         按 **3 段折线** 插值：节点 (0, 1.0) → (1/3, 1 − 0.45·t) →
 *                         (2/3, 1 − 0.78·t) → (1, 1 − t)，t = fTaperPct ÷ 100。
 *                         折线前段缓、后段陡：小卷径段张力衰减慢（防松卷），大卷径段衰减快
 *                         （防内层压溃），与线性锥度件（FB_DL_WinderTensionTaperCtrl）
 *                         的区别即在此曲线形状。
 *                         **卷径有效性闸**：fRollDia ≤ 0 或 > fDiaMax → eFault 且 fTensionOut := 0
 *                         （安全侧直接撤张力，不保留末值）。
 *                         **bEnable = FALSE 语义（R191 二选一，本件选「冻结保持末值」）**：
 *                         张力环的硬切断由上级安全回路负责，本件失能时保持末值不突变。
 * 接口     (Interface)  : 输入 bEnable / bReset / fRollDia / fDiaCore / fDiaMax / fTensionIn /
 *                         fTaperPct / fTensionMin / fTensionMax；输出 fTensionOut（限幅后）/
 *                         fTaperFactor / fDiaRatio / eState / bError / eCause / bValid。
 * 状态迁移表 (State Transition Table)：
 *   ① eIdle → eRun：bEnable 上升（进入计算相）；拍 N 进入（bEnable）/ 本拍行为：不做计算、
 *      输出保持末值 / 拍 N+1 转出至 eRun。
 *   ② eRun → eFault：组态域闸失败（卷芯径 ≤0 / 卷径上下限倒置 / 张力上下限倒置 /
 *      锥度率越域 0..90 / 任一浮点非有限）或卷径有效性闸失败（≤0 或 > fDiaMax）；
 *      拍 N 进入（判据失败）/ 本拍行为：锁存首因、fTensionOut := 0、fTaperFactor := 0 /
 *      拍 N+1 转出至 eFault（段尾迁移闸）。
 *   ③ eRun → eIdle：bEnable 落 FALSE（失能退出，出口冻结保持）。
 *   ④ eIdle → eFault：段尾迁移闸（锁存位已置）。
 *   ⑤ eFault → eIdle：bReset 上升且 NOT bEnable（复位沿要求先失能，可达性自证 R152：
 *      两引脚外部恒可达）；拍 N 进入（复位沿 + 已失能）/ 本拍行为：清锁存与成因码 /
 *      拍 N+1 转出至 eIdle。
 *   ⑥ ELSE（非法枚举值）→ eFault，成因码 eIllegalState（R6 兜底）。
 * 边界     (Boundary)   : ① 卷径先钳位到 [fDiaCore, fDiaMax] 再算比例（r 结构性落在 [0,1]）。
 *                         ② 折线三段的插值分母均为常量（0.33333、0.33334、0.33333），
 *                            编译期非零，结构性无除零（R4）。
 *                         ③ t = fTaperPct ÷ 100.0，除数为字面常量 100.0（非零）。
 *                         ④ 输出张力钳位到 [fTensionMin, fTensionMax]，上限 / 下限饱和各占
 *                            独立成因成员（R190 归因唯一）。
 *                         ⑤ 浮点同值比较统一容差 DL_TTP_EPS（1E-6），禁 `=`。
 *                         ⑥ 零全局耦合（无 GVL / VAR_EXTERNAL / %I / %Q）。
 * 码表     (Codes)      : 本件不占用全局数字码位（R297 零码位范式）；出口为 BOOL + ENUM，
 *                         enum E_DL_TaperCause 归属本文件（全库唯一属主）。信息级
 *                         eSatHigh / eSatLow 永不置 bError；故障级码锁存回放至 bReset 沿。
 * 分工声明 (Scope)      : 线性锥度 + 斜坡限速件为 FB_DL_WinderTensionTaperCtrl（E_DL_WttState
 *                         属主）；本件只做分段折线曲线与钳位，不做斜坡、不做张力闭环。
 * 归属     (Ownership)  : E_DL_WttState 归属 FB_DL_WinderTensionTaperCtrl.st，本件只引用
 *                         不重声明（R264）；E_DL_TaperCause 归属本文件。
 * 红线自检 (Redline)    : R1 ✓ 零 GVL ｜ R2 ✓ 零 %I/%Q ｜ R3 ✓ 纯 IEC ｜ R4 ✓ 卷径域闸 +
 *                         非有限双判 + 常量除法 + 容差比较 ｜ R5 ✓ 逐行同行双语注释
 *                         R6 ✓ 三态 ENUM + CASE + ELSE ｜ R7 N/A（无定时器/边沿实例）
 *                         R14 ✓ 无 PROPERTY ｜ R8/R9 N/A（无 METHOD）
 * 修订历史 (Revision)   : 2026-11-23  v1.0.0  R78-B3 首版
 * 验收向量 (Acceptance) :
 *   V1 fRollDia=100, fDiaCore=100, fDiaMax=800, fTensionIn=50, fTaperPct=30 →
 *      r=0 → k=1.0 → fTensionOut=50.0, bValid=TRUE, eCause=eNone。
 *   V2 其余引脚取 V1 值、fRollDia=333.3 → r≈0.3333 → k=1−0.3×0.45=0.865 → fTensionOut≈43.25（容差 1E-3）。
 *   V3 其余引脚取 V1 值、fRollDia=800 → r=1 → k=0.7 → fTensionOut=35.0。
 *   V4 fRollDia=0.0 → eState=eFault, eCause=eBadDiameter, fTensionOut=0.0, bError=TRUE；
 *      bReset 上升且 bEnable=FALSE → 回 eIdle。
 *   V5 fTaperPct=95（越域）→ eState=eFault, eCause=eBadTaper, fTensionOut=0.0。
 *   V6 fTensionOut 计算得 5.0 而 fTensionMin=10.0 → fTensionOut=10.0, eCause=eSatLow（信息级）。
 *============================================================================*)

(*-----------------------------------------------------------------------------
 * 枚举: E_DL_TaperCause（锥度张力成因码；信息级 = 0..9，故障级 = 10 起）
 *----------------------------------------------------------------------------*)
TYPE E_DL_TaperCause :
(
    eNone         := 0,   // 信息级：计算正常 / Info: computation normal
    eSatHigh      := 1,   // 信息级：输出张力已饱和到上限 / Info: output saturated at the high limit
    eSatLow       := 2,   // 信息级：输出张力已饱和到下限 / Info: output saturated at the low limit
    eBadDiameter  := 10,  // 故障级：卷径反馈无效（≤0 或 > fDiaMax）/ Fault: invalid roll diameter
    eBadConfig    := 11,  // 故障级：卷芯/限值组态倒置或越界 / Fault: inverted or out-of-range configuration
    eBadTaper     := 12,  // 故障级：锥度率越域（0..90）/ Fault: taper percentage out of the 0..90 domain
    eNonFinite    := 13,  // 故障级：入参非有限 / Fault: non-finite input
    eIllegalState := 14   // 故障级：非法状态枚举值 / Fault: illegal state enum value
);
END_TYPE

FUNCTION_BLOCK FB_DL_WinderTensionTaperCalc
VAR_INPUT
    bEnable     : BOOL := FALSE;      // 使能：FALSE 冻结保持末值（本件语义声明）/ Enable, FALSE freezes the last output
    bReset      : BOOL := FALSE;      // 复位（上升沿，需同时 bEnable=FALSE）/ Reset rising edge, requires disabled state
    fRollDia    : REAL := 100.0;      // 当前卷径反馈，有效域 (0, fDiaMax] [mm] / Current roll diameter feedback [mm]
    fDiaCore    : REAL := 100.0;      // 卷芯直径（锥度曲线起点），域 > 0 [mm] / Core diameter, curve origin [mm]
    fDiaMax     : REAL := 800.0;      // 满卷直径（锥度曲线终点），域 > fDiaCore [mm] / Full roll diameter, curve end [mm]
    fTensionIn  : REAL := 50.0;       // 内圈基础张力给定 [N] / Base (inner) tension setpoint [N]
    fTaperPct   : REAL := 30.0;       // 满卷处张力衰减百分比，有效域 0..90 [%] / Tension taper at full roll, domain 0..90 [%]
    fTensionMin : REAL := 0.0;        // 张力输出下限，域 ≥ 0 [N] / Tension output low limit [N]
    fTensionMax : REAL := 200.0;      // 张力输出上限，域 > fTensionMin [N] / Tension output high limit [N]
END_VAR
VAR_OUTPUT
    fTensionOut  : REAL := 0.0;        // 锥度张力输出（限幅后）[N] / Tapered tension output after clamping [N]
    fTaperFactor : REAL := 0.0;        // 本拍锥度系数 k（0..1）[-] / Taper factor k of this scan
    fDiaRatio    : REAL := 0.0;        // 本拍归一化卷径比例 r（0..1）[-] / Normalised diameter ratio r of this scan
    eState       : E_DL_WttState;      // 状态出口（段尾单点映射，引用属主枚举）[-] / State outlet mapped at the tail
    bError       : BOOL;               // 故障锁存标志 [-] / Fault latch flag
    eCause       : E_DL_TaperCause;    // 成因码出口（故障期锁存回放）[-] / Cause code outlet, latched replay
    bValid       : BOOL;               // 张力输出有效回执 [-] / Tension output validity receipt
END_VAR
VAR
    _eState      : E_DL_WttState := E_DL_WttState.eIdle;    // 内部相位（CASE 唯一写入目标）[-] / Internal phase
    _bFaultLatch : BOOL := FALSE;                           // 故障锁存位（仅 bReset 沿清除）[-] / Fault latch bit
    _eCauseLatch : E_DL_TaperCause := E_DL_TaperCause.eNone; // 锁存成因码（FB33-1 锁存回放）[-] / Latched cause code
    _eCauseTmp   : E_DL_TaperCause := E_DL_TaperCause.eNone; // 本拍首个成因（未锁存）[-] / First cause of this scan
    _bCfgOk      : BOOL := TRUE;                            // 组态与入参闸通过标志 [-] / Configuration gate flag
    _fDiaClamped : REAL := 0.0;                             // 钳位后的卷径 [mm] / Clamped roll diameter
    _fRatio       : REAL := 0.0;                            // 归一化卷径比例 r [-] / Normalised diameter ratio
    _fTaperFrac  : REAL := 0.0;                             // 锥度小数 t = fTaperPct/100 [-] / Taper fraction
    _fK1         : REAL := 0.0;                             // 折线节点 1/3 处系数 [-] / Factor at the one-third knot
    _fK2         : REAL := 0.0;                             // 折线节点 2/3 处系数 [-] / Factor at the two-thirds knot
    _fK3         : REAL := 0.0;                             // 折线节点 1 处系数 (1 − t) [-] / Factor at the full-roll knot
    _fK          : REAL := 0.0;                             // 本拍锥度系数 k [-] / Taper factor of this scan
    _fTension     : REAL := 0.0;                            // 钳位前张力 [N] / Tension before clamping
    nSeg         : INT := 0;                                // 折线段号 [1..3] / Piecewise segment index
END_VAR
VAR CONSTANT
    DL_TTP_ZERO  : REAL := 0.0;        // 零基准 [-] / Zero base
    DL_TTP_ONE   : REAL := 1.0;        // 一基准（单位 / 比例上端）[-] / Unity base
    DL_TTP_FULL  : REAL := 100.0;      // 百分比换算分母（非零常量）/ Percentage denominator, a non-zero constant
    DL_TTP_R1    : REAL := 0.33333;    // 折线第 1 节点比例 [-] / First knot ratio
    DL_TTP_R2    : REAL := 0.66667;    // 折线第 2 节点比例 [-] / Second knot ratio
    DL_TTP_KT1   : REAL := 0.45;       // 第 1 节点处衰减占比（占 t 的比例）[-] / Decay share at the first knot
    DL_TTP_KT2   : REAL := 0.78;       // 第 2 节点处衰减占比（占 t 的比例）[-] / Decay share at the second knot
    DL_TTP_D1    : REAL := 0.33333;    // 第 1 段插值分母（R1 − 0）[-] / Denominator of segment one
    DL_TTP_D2    : REAL := 0.33334;    // 第 2 段插值分母（R2 − R1）[-] / Denominator of segment two
    DL_TTP_D3    : REAL := 0.33333;    // 第 3 段插值分母（1 − R2）[-] / Denominator of segment three
    DL_TTP_TPMAX : REAL := 90.0;       // 锥度率上限（> 90% 的衰减无工程意义）[%] / Upper taper limit [%]
    DL_TTP_EPS   : REAL := 1.0E-6;     // 浮点同值比较容差 [-] / Float equality tolerance
END_VAR

(* —— 段 1：当拍工作量预置（单拍标志与中间量，不清锁存/保持量） —— *)
_bCfgOk    := TRUE;                                     // 闸通过标志复位 / Gate flag reset
_eCauseTmp := E_DL_TaperCause.eNone;                     // 当拍成因复位 / Scan cause reset

(* —— 段 2：状态机主体（唯一相位写入点） —— *)
CASE _eState OF
    E_DL_WttState.eIdle :
        IF bEnable THEN
            _eState := E_DL_WttState.eRun;               // 迁移①：进入计算相 / Move to the run phase
        END_IF

    E_DL_WttState.eRun :
        IF NOT bEnable THEN
            _eState := E_DL_WttState.eIdle;              // 迁移③：失能退出（冻结保持）/ Disable exit
        ELSE
            (* —— 段 3：入参非有限闸（R272 全量枚举九个浮点引脚） —— *)
            IF (fRollDia <> fRollDia) OR ((fRollDia - fRollDia) <> DL_TTP_ZERO)
                OR (fDiaCore <> fDiaCore) OR ((fDiaCore - fDiaCore) <> DL_TTP_ZERO)
                OR (fDiaMax <> fDiaMax) OR ((fDiaMax - fDiaMax) <> DL_TTP_ZERO)
                OR (fTensionIn <> fTensionIn) OR ((fTensionIn - fTensionIn) <> DL_TTP_ZERO)
                OR (fTaperPct <> fTaperPct) OR ((fTaperPct - fTaperPct) <> DL_TTP_ZERO)
                OR (fTensionMin <> fTensionMin) OR ((fTensionMin - fTensionMin) <> DL_TTP_ZERO)
                OR (fTensionMax <> fTensionMax) OR ((fTensionMax - fTensionMax) <> DL_TTP_ZERO) THEN
                _bCfgOk    := FALSE;
                _eCauseTmp := E_DL_TaperCause.eNonFinite;    // 故障级：非有限 / Fault: non-finite
            END_IF
            (* —— 段 4：组态域闸（两两倒置 / 越界各自独立成因） —— *)
            IF _bCfgOk THEN
                IF (fDiaCore <= DL_TTP_ZERO) OR (fDiaMax <= fDiaCore) THEN
                    _bCfgOk    := FALSE;
                    _eCauseTmp := E_DL_TaperCause.eBadConfig;      // 故障级：卷径组态倒置
                ELSIF (fTensionMin < DL_TTP_ZERO) OR (fTensionMax <= fTensionMin) THEN
                    _bCfgOk    := FALSE;
                    _eCauseTmp := E_DL_TaperCause.eBadConfig;      // 故障级：张力组态倒置
                ELSIF (fTaperPct < DL_TTP_ZERO) OR (fTaperPct > DL_TTP_TPMAX) THEN
                    _bCfgOk    := FALSE;
                    _eCauseTmp := E_DL_TaperCause.eBadTaper;       // 故障级：锥度率越域
                END_IF
            END_IF
            (* —— 段 5：卷径有效性闸（≤0 或 > 满卷径 → 撤张力） —— *)
            IF _bCfgOk THEN
                IF (fRollDia <= DL_TTP_ZERO) OR (fRollDia > (fDiaMax + DL_TTP_EPS)) THEN
                    _bCfgOk    := FALSE;
                    _eCauseTmp := E_DL_TaperCause.eBadDiameter;    // 故障级：卷径无效
                END_IF
            END_IF

            IF NOT _bCfgOk THEN
                (* 迁移②：锁存首因 + 安全侧撤张力（不保留末值） *)
                _eCauseLatch := _eCauseTmp;                    // 锁存成因 / Latch the cause
                _bFaultLatch := TRUE;                          // 置故障锁存 / Latch the fault
                fTensionOut  := DL_TTP_ZERO;                   // 安全侧：张力输出 0 / Safe side: zero tension
                fTaperFactor := DL_TTP_ZERO;                   // 锥度系数同步清零 / Taper factor zeroed
                _eState      := E_DL_WttState.eFault;          // 迁入故障相 / Move to the fault phase
            ELSE
                (* —— 段 6：比例与三段折线（分母全为编译期非零常量） —— *)
                _fDiaClamped := MIN(MAX(fRollDia, fDiaCore), fDiaMax);         // 卷径先钳位（R4）/ Clamp the diameter first
                _fRatio      := (_fDiaClamped - fDiaCore) / (fDiaMax - fDiaCore);   // 归一化比例 r / Normalised ratio
                _fRatio      := MIN(MAX(_fRatio, DL_TTP_ZERO), DL_TTP_ONE);    // 比例钳到 [0,1] / Clamp the ratio
                _fTaperFrac  := fTaperPct / DL_TTP_FULL;                        // 锥度小数 t / Taper fraction
                _fK1         := DL_TTP_ONE - (_fTaperFrac * DL_TTP_KT1);        // 节点 1/3 系数 / Factor at knot one
                _fK2         := DL_TTP_ONE - (_fTaperFrac * DL_TTP_KT2);        // 节点 2/3 系数 / Factor at knot two
                _fK3         := DL_TTP_ONE - _fTaperFrac;                       // 满卷节点系数 / Factor at full roll
                IF _fRatio <= DL_TTP_R1 THEN
                    nSeg := 1;                                                  // 第 1 段 / Segment one
                ELSIF _fRatio <= DL_TTP_R2 THEN
                    nSeg := 2;                                                  // 第 2 段 / Segment two
                ELSE
                    nSeg := 3;                                                  // 第 3 段 / Segment three
                END_IF
                CASE nSeg OF
                    1 :
                        _fK := DL_TTP_ONE + ((_fK1 - DL_TTP_ONE) * (_fRatio / DL_TTP_D1));      // 段 1 线性插值
                    2 :
                        _fK := _fK1 + ((_fK2 - _fK1) * ((_fRatio - DL_TTP_R1) / DL_TTP_D2));    // 段 2 线性插值
                    3 :
                        _fK := _fK2 + ((_fK3 - _fK2) * ((_fRatio - DL_TTP_R2) / DL_TTP_D3));    // 段 3 线性插值
                ELSE
                    _fK := DL_TTP_ONE;                                          // 兜底：恒张力系数 / Fallback: constant factor
                END_CASE
                _fTension := fTensionIn * _fK;                                   // 锥度张力 = 基础张力 × k / Tapered tension
                (* —— 段 7：输出钳位（上/下限独立成因，R190） —— *)
                IF _fTension > fTensionMax THEN
                    fTensionOut := fTensionMax;                                  // 上限饱和 / Saturate high
                    eCause      := E_DL_TaperCause.eSatHigh;                     // 信息级：上限饱和 / Info: saturated high
                ELSIF _fTension < fTensionMin THEN
                    fTensionOut := fTensionMin;                                  // 下限饱和 / Saturate low
                    eCause      := E_DL_TaperCause.eSatLow;                      // 信息级：下限饱和 / Info: saturated low
                ELSE
                    fTensionOut := _fTension;                                    // 限内直通 / Pass-through
                    eCause      := E_DL_TaperCause.eNone;                        // 信息级：正常 / Info: normal
                END_IF
                fTaperFactor := _fK;                                             // 锥度系数出口 / Taper factor outlet
                fDiaRatio    := _fRatio;                                         // 卷径比例出口 / Diameter ratio outlet
            END_IF
        END_IF

    E_DL_WttState.eFault :
        (* 迁移⑤：唯一出口 —— bReset 沿 + 已失能 *)
        IF bReset AND (NOT bEnable) THEN
            _bFaultLatch := FALSE;                             // 清故障锁存 / Clear the latch
            _eCauseLatch := E_DL_TaperCause.eNone;             // 清锁存成因 / Clear the latched cause
            eCause       := E_DL_TaperCause.eNone;             // 出口同步归零 / Outlet follows
            _eState      := E_DL_WttState.eIdle;               // 回空闲相 / Back to idle
        END_IF

ELSE
    (* 迁移⑥：非法枚举兜底（R6） *)
    _eCauseLatch := E_DL_TaperCause.eIllegalState;             // 故障级：非法状态
    _bFaultLatch := TRUE;                                      // 置锁存 / Latch
    fTensionOut  := DL_TTP_ZERO;                               // 安全侧撤张力 / Safe side: zero tension
    _eState      := E_DL_WttState.eFault;                      // 迁入故障相 / Move to fault
END_CASE

(* —— 段 8：段尾故障迁移闸（锁存与迁相分离，FB50-1④） —— *)
IF _bFaultLatch AND (_eState <> E_DL_WttState.eFault) THEN
    _eState := E_DL_WttState.eFault;                           // 锁存即迁相 / Latch forces the fault phase
END_IF

(* —— 段 9：统一出口（状态映射 + 锁存回放） —— *)
eState := _eState;                                             // 相位映射 / Phase mapping
bError := _bFaultLatch;                                        // 故障标志取锁存位 / Fault flag from the latch
IF _bFaultLatch THEN
    eCause := _eCauseLatch;                                    // 故障期回放锁存码（FB33-1）/ Replay the latched code
END_IF
bValid := (_eState = E_DL_WttState.eRun) AND (NOT _bFaultLatch);   // 仅计算相且无锁存时有效 / Valid only in run without a latch
END_FUNCTION_BLOCK
